// TIA Portal V21 export
// export: Created 2026-11-07T15:50:51.3358476Z, ExportSetting WithDefaults, DisplayName Totally Integrated Automation Portal, DisplayVersion V21, DisplayName STEP 7 Professional, DisplayVersion V21, DisplayName STEP 7 Safety, DisplayVersion V21, DisplayName Tech WebApplication, DisplayVersion V21, DisplayName WinCC Basic/Comfort/Advanced, DisplayVersion V21, DisplayName WinCC Unified, DisplayVersion V21
Screen "R07_MoveV"  1024x768, Number=47, Template=Tpl
  ScreenLayer 
    Rectangle "P_CraneY" at 10,10 size 100x30  StyleItem=Rectangle
      VerticalMovementAnimation "VerticalMovementAnimation"  RangeEnd=100, YDelta=-10
        tag 
